FUNCTION_BLOCK CompositeHashTest (* Composite FB containing a basic FB *)
  (* Standard: 61499-1; Description: Copyright (c) 2026 Martin Erich Jobst This program and the accompanying materials are made available under the terms of the Eclipse Public License 2.0 which is available at https://www.eclipse.org/legal/epl-2.0/ SPDX-License-Identifier: EPL-2.0 *)
  (* Version 1.0, 2026-10-28, Martin Jobst *)
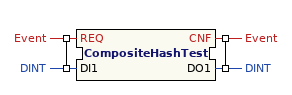
  EVENT_INPUT
    REQ WITH DI1; (* Request *)
  END_EVENT
  EVENT_OUTPUT
    CNF WITH DO1; (* Confirmation *)
  END_EVENT
  VAR_INPUT
    DI1 : DINT := DINT#42;
  END_VAR
  VAR_OUTPUT
    DO1 : DINT;
  END_VAR
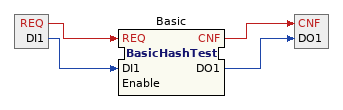
  FBS
    Basic : BasicHashTest;
  END_FBS
  EVENT_CONNECTIONS
    REQ TO Basic.REQ;
    Basic.CNF TO CNF;
  END_CONNECTIONS
  DATA_CONNECTIONS
    DI1 TO Basic.DI1;
    Basic.DO1 TO DO1;
  END_CONNECTIONS
END_FUNCTION_BLOCK
